(* IEC 61131-3 sources: TrakMap/InstallerSetup/Installer AS Technology Solution/Logical/Libraries/snprintf, 3 files *)

(* ---- snprintf.typ ---- *)
(********************************************************************
 * COPYRIGHT -- B&R
 ********************************************************************
 * Library: snprintf
 * File: snprintf.typ
 * Author: buchananw
 * Created: April 15, 2009
 ********************************************************************
 * Data types of library snprintf
 ********************************************************************)

TYPE

END_TYPE

(* ---- snprintf.fun ---- *)
(********************************************************************
 * COPYRIGHT -- B&R
 ********************************************************************
 * Library: snprintf
 * File: snprintf.fun
 * Author: buchananw
 * Created: April 15, 2009
 ********************************************************************
 * Functions and function blocks of library snprintf
 ********************************************************************)

FUNCTION snprintf2 : SINT
END_FUNCTION

(* ---- snprintf.var ---- *)
(********************************************************************
 * COPYRIGHT -- B&R
 ********************************************************************
 * Library: snprintf
 * File: snprintf.var
 * Author: buchananw
 * Created: April 15, 2009
 ********************************************************************
 * Constants of library snprintf
 ********************************************************************)

VAR CONSTANT

END_VAR
